{attribute 'TcHmiSymbol.ShowRecursively'}
TYPE T_NOTT_DETECTOR_POWER_STAT :
STRUCT
    bPowerOn: BOOL;
    bCurrentValid: BOOL;
    bMeasurementStale: BOOL;
    bUnderrange: BOOL;
    bOverrange: BOOL;
    bExtendedRange: BOOL;
    bDataInvalid: BOOL;
    bRangeInvalid: BOOL;
    bAutorangeDisabled: BOOL;
    bConversionError: BOOL;
    bCalibrating: BOOL;
    bPdoInvalid: BOOL;
    bPdoToggle: BOOL;
    bMeterOperational: BOOL;
    bFuseOperational: BOOL;
    bConfigValid: BOOL;
    bOvercurrentTrip: BOOL;
    bShutdownUnconfirmed: BOOL;
    bPermitOn: BOOL;
    bPermitTripReset: BOOL;
    bAlarm: BOOL;
    bWarning: BOOL;
    lrCurrent_A: LREAL;
    lrTripCurrent_A: LREAL;
    nMeterStatus: UINT;
    nLastCommand: DINT;
    sStatus: STRING(255);
    sCommandResult: STRING(255);
    sMeasurementStatus: STRING(255);
END_STRUCT
END_TYPE

(* stored: Version 1.1.0.1, ProductVersion 3.1.4026.20
   DUT T_NOTT_DETECTOR_POWER_STAT: Id {6ddfe093-2ee4-49bf-a222-2570d444108a} *)
